FUNCTION "FRK_PersistDirty" : Void
{ S7_Optimized_Access := 'TRUE' }
VERSION : 0.1
VAR_INPUT
    Slot : Int;
END_VAR
VAR_TEMP
    Stamp : LDT;
    NativeResult : Int;
END_VAR
BEGIN
    IF #Slot < 1 OR #Slot > 12 THEN RETURN; END_IF;
    IF NOT "FRK_PersistConsumers".Rows[#Slot].Dirty THEN
        #NativeResult := RD_SYS_T(OUT => #Stamp);
        IF "FRK_PersistConsumers".Rows[#Slot].Ticket = 0 THEN "FRK_PersistConsumers".Rows[#Slot].PendingSince := #Stamp;
        ELSE "FRK_PersistConsumers".Rows[#Slot].NextSince := #Stamp; END_IF;
    END_IF;
    "FRK_PersistConsumers".Rows[#Slot].Dirty := TRUE;
END_FUNCTION
FUNCTION "FRK_PersistConfigSlot" : Int
{ S7_Optimized_Access := 'TRUE' }
VERSION : 0.1
VAR_INPUT
    Scope : String;
    ModelCode : String;
    Kind : DInt;
END_VAR
BEGIN
    #FRK_PersistConfigSlot := 0;
    IF #Scope = 'PressDemo' AND #ModelCode = '' AND #Kind = 1 THEN #FRK_PersistConfigSlot := 1; RETURN; END_IF;
    IF #Scope = 'PressDemo' AND #ModelCode = '' AND #Kind = 1 THEN #FRK_PersistConfigSlot := 1; RETURN; END_IF;
    IF #Scope = 'PressDemo' AND #ModelCode = 'ALUMINUM' AND #Kind = 0 THEN #FRK_PersistConfigSlot := 2; RETURN; END_IF;
    IF #Scope = 'PressDemo' AND #ModelCode = 'ALUMINUM' AND #Kind = 0 THEN #FRK_PersistConfigSlot := 2; RETURN; END_IF;
    IF #Scope = 'PressDemo' AND #ModelCode = 'ALUMINUM' AND #Kind = 0 THEN #FRK_PersistConfigSlot := 2; RETURN; END_IF;
    IF #Scope = 'PressDemo' AND #ModelCode = 'ALUMINUM' AND #Kind = 0 THEN #FRK_PersistConfigSlot := 2; RETURN; END_IF;
    IF #Scope = 'PressDemo' AND #ModelCode = 'ALUMINUM' AND #Kind = 0 THEN #FRK_PersistConfigSlot := 2; RETURN; END_IF;
    IF #Scope = 'PressDemo' AND #ModelCode = 'PLASTIC' AND #Kind = 0 THEN #FRK_PersistConfigSlot := 3; RETURN; END_IF;
    IF #Scope = 'PressDemo' AND #ModelCode = 'PLASTIC' AND #Kind = 0 THEN #FRK_PersistConfigSlot := 3; RETURN; END_IF;
    IF #Scope = 'PressDemo' AND #ModelCode = 'PLASTIC' AND #Kind = 0 THEN #FRK_PersistConfigSlot := 3; RETURN; END_IF;
    IF #Scope = 'PressDemo' AND #ModelCode = 'PLASTIC' AND #Kind = 0 THEN #FRK_PersistConfigSlot := 3; RETURN; END_IF;
    IF #Scope = 'PressDemo' AND #ModelCode = 'PLASTIC' AND #Kind = 0 THEN #FRK_PersistConfigSlot := 3; RETURN; END_IF;
    IF #Scope = 'PressDemo' AND #ModelCode = 'STEEL' AND #Kind = 0 THEN #FRK_PersistConfigSlot := 4; RETURN; END_IF;
    IF #Scope = 'PressDemo' AND #ModelCode = 'STEEL' AND #Kind = 0 THEN #FRK_PersistConfigSlot := 4; RETURN; END_IF;
    IF #Scope = 'PressDemo' AND #ModelCode = 'STEEL' AND #Kind = 0 THEN #FRK_PersistConfigSlot := 4; RETURN; END_IF;
    IF #Scope = 'PressDemo' AND #ModelCode = 'STEEL' AND #Kind = 0 THEN #FRK_PersistConfigSlot := 4; RETURN; END_IF;
    IF #Scope = 'PressDemo' AND #ModelCode = 'STEEL' AND #Kind = 0 THEN #FRK_PersistConfigSlot := 4; RETURN; END_IF;
    IF #Kind = 0 AND (#Scope = 'PressDemo') THEN #FRK_PersistConfigSlot := 12; RETURN; END_IF;
END_FUNCTION
FUNCTION "FRK_PersistUsersDirty" : Void
{ S7_Optimized_Access := 'TRUE' }
VERSION : 0.1
BEGIN
    "FRK_PersistDirty"(Slot := 10);
END_FUNCTION
FUNCTION "FRK_PersistPolicyDirty" : Void
{ S7_Optimized_Access := 'TRUE' }
VERSION : 0.1
VAR_INPUT
    RootIndex : Int;
END_VAR
BEGIN
    IF #RootIndex = 1 THEN "FRK_PersistDirty"(Slot := 5); END_IF;
END_FUNCTION
FUNCTION "FRK_PersistSetDirty" : Void
{ S7_Optimized_Access := 'TRUE' }
VERSION : 0.1
VAR_INPUT
    RootIndex : Int;
    Ordinal : Int;
END_VAR
BEGIN
    IF #RootIndex = 1 AND #Ordinal = 1 THEN "FRK_PersistDirty"(Slot := 6); END_IF;
    IF #RootIndex = 1 AND #Ordinal = 2 THEN "FRK_PersistDirty"(Slot := 7); END_IF;
    IF #RootIndex = 1 AND #Ordinal = 3 THEN "FRK_PersistDirty"(Slot := 8); END_IF;
    IF #RootIndex = 1 AND #Ordinal = 4 THEN "FRK_PersistDirty"(Slot := 9); END_IF;
END_FUNCTION
FUNCTION "FRK_PersistModelDirty" : Void
{ S7_Optimized_Access := 'TRUE' }
VERSION : 0.1
VAR_INPUT
    RootIndex : Int;
END_VAR
BEGIN
    IF #RootIndex = 1 THEN "FRK_PersistDirty"(Slot := 1); END_IF;
END_FUNCTION
FUNCTION "FRK_PersistModelsDirty" : Void
{ S7_Optimized_Access := 'TRUE' }
VERSION : 0.1
VAR_INPUT
    RootIndex : Int;
END_VAR
BEGIN
    IF #RootIndex = 1 THEN "FRK_PersistDirty"(Slot := 12); END_IF;
END_FUNCTION
FUNCTION "FRK_PersistModelsSaved" : Bool
{ S7_Optimized_Access := 'TRUE' }
VERSION : 0.1
VAR_INPUT
    RootIndex : Int;
END_VAR
BEGIN
    #FRK_PersistModelsSaved := FALSE;
    IF NOT "FRK_PersistConsumers".Ready THEN RETURN; END_IF;
    IF #RootIndex = 1 THEN
        #FRK_PersistModelsSaved := "FRK_PersistConsumers".Rows[12].State = 2 AND "FRK_PersistConsumers".Rows[12].Ticket = 0 AND NOT "FRK_PersistConsumers".Rows[12].Dirty AND NOT "FRK_PersistConsumers".Rows[12].Failed AND (NOT "FRK_PersistConsumers".Rows[12].Rejected OR "FRK_PersistConsumers".Rows[12].Acknowledged);
    END_IF;
END_FUNCTION
FUNCTION "FRK_PersistVirginConfig" : Bool
{ S7_Optimized_Access := 'TRUE' }
VERSION : 0.1
VAR_INPUT
    Scope : String;
    ModelCode : String;
    Kind : DInt;
END_VAR
VAR_TEMP
    Slot : Int;
END_VAR
BEGIN
    #FRK_PersistVirginConfig := FALSE;
    #Slot := "FRK_PersistConfigSlot"(Scope := #Scope, ModelCode := #ModelCode, Kind := #Kind);
    IF #Slot > 0 THEN #FRK_PersistVirginConfig := "FRK_PersistConsumers".Rows[#Slot].Virgin; END_IF;
END_FUNCTION
FUNCTION "FRK_PersistLineTick" : Void
{ S7_Optimized_Access := 'TRUE' }
VERSION : 0.1
BEGIN
    IF "FRK_PersistConsumers".Ready AND "FRK_Line".Data.Dirty THEN
        "FRK_PersistDirty"(Slot := 11);
        "FRK_Line".Data.Dirty := FALSE;
    END_IF;
END_FUNCTION
